{attribute 'qualified_only'}
VAR_GLOBAL
	AbsoluteBetaPosition AT %I* : DINT;
	AbsoluteLinearPosition AT %I* : DINT;
	AbsoluteTetaPosition AT %I* : DINT;
END_VAR

(* stored: Version 1.1.0.1, ProductVersion 3.1.4024.15
   GVL GVL_AbsoluteEncoders: Id {41acc025-99db-4313-b396-7394fb224741} *)
